Fanuc KAREL source: KO00047.KL

PROGRAM KO00047
%NOLOCKGROUP
%ENVIRONMENT MIR
VAR
  P1: POSITION
  P2: JOINTPOS
  F: BOOLEAN
  OUT: XYZWPREXT
BEGIN
  F = TRUE
  OUT = MIRROR(P1, P2, F)
END KO00047
